FUNCTION_BLOCK FB_GCodeUSB EXTENDS FB_RecipeBase

METHOD Build : BOOL
VAR
      i          : INT;
END_VAR

VAR_INST
    nBuildStep : INT;
    machineConfig : ST_GantryXYZ_Config;
END_VAR
_Done := FALSE;
_Error := FALSE;

IF LEN(_Config.GCodePath) > 0 THEN
    _Config.IsValid := TRUE;
    _Done           := TRUE;
    Build           := TRUE;
ELSE
    _Config.IsValid := FALSE;
    _Error          := TRUE;
    Build           := FALSE;
END_IF
END_METHOD

PROPERTY ExecutionRoute : E_ExecutionRoute
GET
ExecutionRoute := E_ExecutionRoute.eGCode;
END_GET
END_PROPERTY

END_FUNCTION_BLOCK

(* stored: Version 1.1.0.1, ProductVersion 3.1.4024.15
   POU FB_GCodeUSB: Id {fccba36f-1e04-4dd4-8f5d-37009967fb17}, SpecialFunc None
   Method Build: Id {a9c31ce6-ed3e-43ff-bafc-85dc97fdd881}
   Property ExecutionRoute: Id {e6277044-3ac9-41ce-80fb-2e38121afadb}
   Get Get: Id {077466b1-15fc-433c-99bc-d5b5661032e0} *)
